RoboDK station: hand_motion - Contactile.rdk

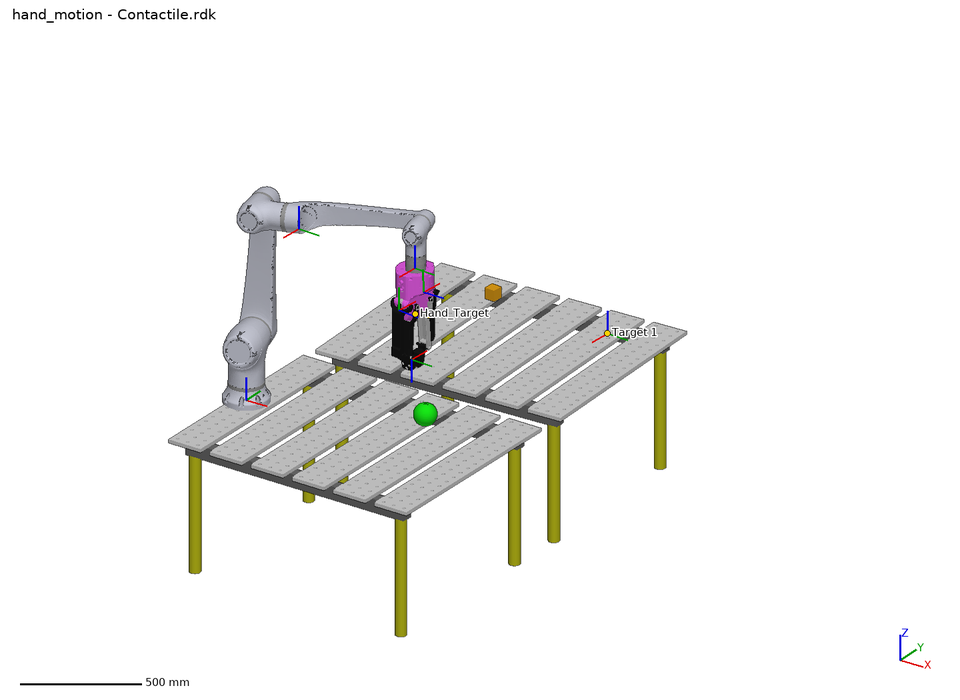
[picture v0: the station drawn from its stored meshes, robots at their saved joint values, targets as dots, program paths as lines]
Station hand_motion - Contactile (saved by RoboDK 6.0.6). Poses are relative to the parent item; angles as X-Y-Z fixed-axis rotations.
  - frame Neura LARA 8 Base at (0, 0, 0) mm
    - robot Neura LARA 8: 6 axes
        modified DH rows (alpha deg, a mm, theta deg, d mm): 0, 0, 0, 260; -90, 0, -90, 0; 0, 600, -90, 0; -90, 0, 0, 700; 90, 0, 0, 0; -90, 0, 180, 179.5
        joint limits [-180, -135, -155, -180, -180, -360] to [180, 135, 155, 180, 180, 360]; home [0, 0, 90, 0, 90, 0]; saved at [15.447, 3.692, 83.427, -0.003, 92.872, 108.157]
      - tool GAL2_B1.1_CustomerFacing_88mm, TCP at (0, 0, 200) mm, size 76 x 196.6 x 204.3 mm, geometry from GAL2_B1.1_CustomerFacing_88mm.STEP
      - frame Contactile_Gripper_Mount at (10.68, -612.07, -1.87) mm, rotated rx -180 ry 0 rz 180 deg
        - frame GAL2_MASTER Base at (0, 1600, 0) mm
          - robot GAL2_MASTER: 1 axes
              modified DH rows (alpha deg, a mm, theta deg, d mm): 0, 0, 0, 0
              joint limits [0] to [60]; home [0]; saved at [0]
          - target Target 1 (Cartesian target) at (0, 0, 0) mm; joints [0]
          - target Target 2 (Cartesian target) at (0, 0, 0) mm, rotated rx 0 ry 0 rz 6.07 deg; joints [6.07]
        - object link2 at (-84.12, -356.94, -128.79) mm, rotated rx 89.64 ry -0.03 rz -180 deg, size 53 x 255.4 x 102.9 mm, geometry from link2.STL
        - object link1 at (77.57, -359.17, -129.31) mm, rotated rx 179.86 ry -2.12 rz 89.36 deg, size 102.9 x 53 x 255.4 mm, geometry from link1.STL
        - object coupler2 at (-45, -441.52, -148.1) mm, rotated rx 90 ry 9.72 rz 0 deg, size 42.5 x 255.4 x 102.9 mm, geometry from coupler2.STL
        - object coupler1 at (42.87, -442.73, -146.97) mm, rotated rx -90.24 ry 7.58 rz 178.05 deg, size 42.5 x 255.4 x 102.9 mm, geometry from coupler1.STL
        - object base_link at (0, -400, 0) mm, size 203.2 x 159.6 x 215 mm, geometry from base_link.STL
        - Python program Controller (listed below)
        - frame coupler1_mech Base at (0, 600, 0) mm
          - robot coupler1_mech: 1 axes
              modified DH rows (alpha deg, a mm, theta deg, d mm): 0, 0, 0, 0
              base shift (42.87, -442.73, -146.97) mm, rotated rx -90.24 ry 7.58 rz 178.05 deg
              joint limits [-90] to [90]; home [0]; saved at [0]
        - frame coupler2_mech Base at (0, 600, 0) mm
          - robot coupler2_mech: 1 axes
              modified DH rows (alpha deg, a mm, theta deg, d mm): 0, 0, 0, 0
              base shift (-45, -441.52, -148.1) mm, rotated rx 90 ry 9.72 rz 0 deg
              joint limits [-90] to [90]; home [0]; saved at [0]
        - frame link2_mech Base at (-78.92, 585.58, -145.76) mm, rotated rx 88.15 ry -0.03 rz 179.02 deg
          - robot link2_mech: 1 axes
              modified DH rows (alpha deg, a mm, theta deg, d mm): 0, 0, 0, 0
              joint limits [-90] to [90]; home [0]; saved at [0]
        - frame link1_mech Base at (97.92, 593.2, -156.32) mm, rotated rx 90.19 ry 0.13 rz 176.76 deg
          - robot link1_mech: 1 axes
              modified DH rows (alpha deg, a mm, theta deg, d mm): 0, 0, 0, 0
              joint limits [-90] to [90]; home [0]; saved at [0]
        - Python program GAL2_V2 (listed below)
      - frame Grip_Attach_Frame at (0, -20.7, 414.56) mm
    - target Hand_Target (Cartesian target) at (711.17, 196.5, 514.44) mm, rotated rx 179.99 ry 0 rz 87.29 deg; joints [-2.712, 0.991, 79.111, 0, 99.898, -2.712] of Neura LARA 8
    - target Hand_Taught_Target_001 (Cartesian target) at (761.71, 216.75, 515.25) mm, rotated rx 179.99 ry 0 rz 87.29 deg; joints [15.886, 8.932, 77.627, -0.003, 93.432, 108.595] of Neura LARA 8
    - object Sphere D100mm at (744.71, 217.15, 58.5) mm, rotated rx 179.99 ry 0 rz 87.29 deg, size 100 x 100 x 100 mm, geometry from Sphere-D100mm.sld
  - object Table 1200x1000mm (Welding) at (543.39, 0, 0) mm, size 1193.8 x 965.2 x 609.6 mm, geometry from Table-1200x1000mm-Welding.sld
  - object Cube 50mm at (0, 0, 0) mm, size 100 x 100 x 100 mm, geometry from Cube-50mm.sld
  - object Table 1200x1000mm (Welding) at (534.06, 1058.97, 0) mm, rotated rx 0 ry 0 rz 2.59 deg, size 1193.8 x 965.2 x 609.6 mm, geometry from Table-1200x1000mm-Welding.sld
  - Python program Prog3 (listed below)

--- Python program Controller ---
from robodk.robolink import *
from robodk.robomath import *
import time

# ------------------------------------------------------------
# Connect to RoboDK
# ------------------------------------------------------------
RDK = Robolink()

# ------------------------------------------------------------
# Mechanism names
# ------------------------------------------------------------
MECHANISMS = {
    'finger1'  : 'finger1_mech',
    'finger2'  : 'finger2_mech',
    'coupler1' : 'coupler1_mech',
    'coupler2' : 'coupler2_mech',
    'link1'    : 'link1_mech',
    'link2'    : 'link2_mech'
}

# ------------------------------------------------------------
# Get mechanism safely
# ------------------------------------------------------------
def get_mech(name):

    mech = RDK.Item(name)

    if not mech.Valid():
        raise Exception('Missing mechanism: ' + name)

    return mech

# ------------------------------------------------------------
# Load all mechanisms
# ------------------------------------------------------------
finger1  = get_mech(MECHANISMS['finger1'])
finger2  = get_mech(MECHANISMS['finger2'])
coupler1 = get_mech(MECHANISMS['coupler1'])
coupler2 = get_mech(MECHANISMS['coupler2'])
link1    = get_mech(MECHANISMS['link1'])
link2    = get_mech(MECHANISMS['link2'])

# ------------------------------------------------------------
# Set one revolute joint value
# ------------------------------------------------------------
def set_joint(mech, value_deg):

    joints = mech.Joints().list()

    joints[0] = value_deg

    mech.setJoints(joints)

# ------------------------------------------------------------
# MASTER CONTACTILE CONTROL FUNCTION
# ------------------------------------------------------------
# opening_deg:
#     0   = fully closed
#     35  = open
#
# IMPORTANT:
# THESE RATIOS ARE ONLY INITIAL ESTIMATES.
#
# YOU MUST CALIBRATE THEM
# AGAINST THE REAL GRIPPER.
# ------------------------------------------------------------
def set_contactile(opening_deg):

    # -----------------------------
    # Main fingers
    # -----------------------------
    set_joint(finger1,  opening_deg)
    set_joint(finger2, -opening_deg)

    # -----------------------------
    # Coupler links
    # -----------------------------
    set_joint(coupler1,  0.60 * opening_deg)
    set_joint(coupler2, -0.60 * opening_deg)

    # -----------------------------
    # Secondary linkage arms
    # -----------------------------
    set_joint(link1,  1.20 * opening_deg)
    set_joint(link2, -1.20 * opening_deg)

# ------------------------------------------------------------
# SIMPLE OPEN/CLOSE TEST
# ------------------------------------------------------------
def animate_gripper():

    # Open
    for i in range(51):

        a = 35.0 * i / 50.0

        set_contactile(a)

        time.sleep(0.02)

    time.sleep(0.5)

    # Close
    for i in range(51):

        a = 35.0 * (1.0 - i / 50.0)

        set_contactile(a)

        time.sleep(0.02)

# ------------------------------------------------------------
# MAIN
# ------------------------------------------------------------
print('Running Contactile synchronization controller...')

animate_gripper()

print('Finished.')

--- Python program GAL2_V2 ---
# ============================================================
# Contactile GAL2 - Script 3
# RoboDK Synchronization Controller
#
# PURPOSE:
# Reads the GAL2_MASTER joint and synchronizes all six
# nested mechanisms according to the URDF mimic relationships.
#
# REQUIREMENTS:
#
# Existing mechanisms:
#   GAL2_MASTER
#   link1_mech
#   finger1_mech
#   coupler1_mech
#   link2_mech
#   finger2_mech
#   coupler2_mech
#
# Run this script once and leave it running.
# Then move the GAL2_MASTER slider.
# ============================================================

from robodk.robolink import *
from robodk.robomath import *
import time

RDK = Robolink()

# ------------------------------------------------------------
# Get mechanism safely
# ------------------------------------------------------------
def get_item(name):
    item = RDK.Item(name)
    if not item.Valid():
        raise Exception("Missing item: " + name)
    return item

# ------------------------------------------------------------
# Mechanisms
# ------------------------------------------------------------
master    = get_item("GAL2_MASTER")

link1     = get_item("link1_mech")

coupler1  = get_item("coupler1_mech")

link2     = get_item("link2_mech")

coupler2  = get_item("coupler2_mech")

# ------------------------------------------------------------
# Helper
# ------------------------------------------------------------
def set_joint(mech, angle):

    joints = mech.Joints().list()

    joints[0] = angle

    mech.setJoints(joints)

# ------------------------------------------------------------
# Main Loop
# ------------------------------------------------------------
print("GAL2 Synchronization Running...")

previous_theta = None

while True:

    theta = master.Joints().list()[0]

    # Only update if the slider moved
    if theta != previous_theta:

        # ----------------------------------------------------
        # URDF Mimic Relationships
        # ----------------------------------------------------

        # Master
        set_joint(link1, -theta)


        # b_to_c1
        set_joint(coupler1, theta)

        # b_to_l2
        set_joint(link2, theta)

        # b_to_c2
        set_joint(coupler2, theta)

        previous_theta = theta

    time.sleep(0.01)

--- Python program Prog3 ---
from robodk.robolink import *
import time

RDK = Robolink()

sphere = RDK.Item("Sphere D100mm")
link1_mech = RDK.Item("link1_mech")
link2_mech = RDK.Item("link2_mech")

if not sphere.Valid():
    raise Exception("Sphere D100mm not found")

if not link1_mech.Valid():
    raise Exception("link1_mech not found")

if not link2_mech.Valid():
    raise Exception("link2_mech not found")

print("Collision test running.")
print("Move GAL2_MASTER slowly toward closed.")

while True:
    left_contact = RDK.Collision(link1_mech, sphere) > 0
    right_contact = RDK.Collision(link2_mech, sphere) > 0

    if left_contact or right_contact:
        # Red when either side touches
        sphere.setColor([1.0, 0.0, 0.0, 1.0])

        RDK.ShowMessage(
            f"CONTACT: Left={left_contact}, Right={right_contact}",
            False,
        )
    else:
        # Green when there is no contact
        sphere.setColor([0.0, 1.0, 0.0, 1.0])

        RDK.ShowMessage(
            "No finger contact",
            False,
        )

    time.sleep(0.05)
